      R_g[4,14] := -0.11583298;
      R_g[4,15] := 0.43668517;
      R_g[5,0] := -0.15006073;
      R_g[5,1] := 0.14857836;
      R_g[5,2] := 0.09219331;
      R_g[5,3] := 0.24307117;
      R_g[5,4] := 0.02014972;
      R_g[5,5] := -1.73904812;
      R_g[5,6] := -0.06327479;
      R_g[5,7] := 0.09475522;
      R_g[5,8] := -0.05716670;
      R_g[5,9] := 0.00648821;
      R_g[5,10] := -0.08605717;
      R_g[5,11] := 0.04396249;
      R_g[5,12] := 0.19865264;
      R_g[5,13] := 0.21015443;
      R_g[5,14] := -0.04510098;
      R_g[5,15] := -0.05707484;
      R_g[6,0] := 0.05463404;
      R_g[6,1] := -0.24671683;
      R_g[6,2] := 0.14945947;
      R_g[6,3] := 0.27781609;
      R_g[6,4] := 0.05857803;
      R_g[6,5] := -0.09827307;
      R_g[6,6] := -1.36955547;
      R_g[6,7] := 0.03997089;
      R_g[6,8] := 0.10697827;
      R_g[6,9] := -0.15282896;
      R_g[6,10] := -0.11458242;
      R_g[6,11] := 0.23231277;
      R_g[6,12] := 0.06463466;
      R_g[6,13] := -0.04114177;
      R_g[6,14] := 0.01473683;
      R_g[6,15] := 0.09800901;
      R_g[7,0] := 0.03089882;
      R_g[7,1] := -0.12866169;
      R_g[7,2] := -0.14488882;
      R_g[7,3] := 0.08099888;
      R_g[7,4] := -0.01760847;
      R_g[7,5] := 0.12323798;
      R_g[7,6] := 0.01051104;
      R_g[7,7] := -1.43148434;
      R_g[7,8] := 0.05538348;
      R_g[7,9] := 0.08765257;
      R_g[7,10] := 0.04525751;
      R_g[7,11] := -0.08530193;
      R_g[7,12] := 0.06940229;
      R_g[7,13] := 0.20471461;
      R_g[7,14] := 0.11143748;
      R_g[7,15] := -0.01617558;
      R_g[8,0] := 0.00375073;
      R_g[8,1] := 0.05561948;
      R_g[8,2] := 0.07504495;
      R_g[8,3] := 0.13846794;
      R_g[8,4] := 0.01292397;
      R_g[8,5] := -0.12762521;
      R_g[8,6] := 0.00967023;
      R_g[8,7] := -0.02755805;
      R_g[8,8] := -1.64812148;
      R_g[8,9] := 0.12763990;
      R_g[8,10] := 0.15346305;
      R_g[8,11] := -0.01111799;
      R_g[8,12] := 0.17867428;
      R_g[8,13] := -0.14499415;
      R_g[8,14] := -0.04605825;
      R_g[8,15] := 0.04006226;
      R_g[9,0] := 0.07299295;
      R_g[9,1] := -0.19717526;
      R_g[9,2] := -0.09354591;
      R_g[9,3] := 0.11423204;
      R_g[9,4] := 0.18770669;
      R_g[9,5] := -0.18770079;
      R_g[9,6] := 0.17637083;
      R_g[9,7] := -0.00016326;
      R_g[9,8] := 0.05343577;
      R_g[9,9] := -1.98581898;
      R_g[9,10] := -0.07635771;
      R_g[9,11] := 0.00779606;
      R_g[9,12] := -0.21436475;
      R_g[9,13] := 0.14591467;
      R_g[9,14] := 0.07554781;
      R_g[9,15] := -0.05975449;
      R_g[10,0] := -0.25483418;
      R_g[10,1] := 0.06535473;
      R_g[10,2] := -0.15168764;
      R_g[10,3] := -0.13676204;
      R_g[10,4] := 0.13715985;
      R_g[10,5] := -0.04971113;
      R_g[10,6] := -0.04342166;
      R_g[10,7] := 0.13203837;
      R_g[10,8] := -0.05174213;
      R_g[10,9] := 0.17224205;
      R_g[10,10] := -1.54585338;
      R_g[10,11] := 0.08824725;
      R_g[10,12] := 0.54317200;
      R_g[10,13] := -0.00582574;
      R_g[10,14] := -0.18427853;
      R_g[10,15] := -0.08446352;
      R_g[11,0] := -0.01310127;
      R_g[11,1] := 0.35428202;
      R_g[11,2] := -0.22564830;
      R_g[11,3] := -0.47703940;
      R_g[11,4] := 0.02761533;
      R_g[11,5] := -0.02962572;
      R_g[11,6] := 0.06179708;
      R_g[11,7] := -0.01533620;
      R_g[11,8] := 0.04956101;
      R_g[11,9] := 0.15626863;
      R_g[11,10] := -0.12132444;
      R_g[11,11] := -0.90700060;
      R_g[11,12] := 0.20753333;
      R_g[11,13] := -0.08345811;
      R_g[11,14] := -0.30101308;
      R_g[11,15] := -0.34388351;
      R_g[12,0] := 0.15464328;
      R_g[12,1] := -0.19553624;
      R_g[12,2] := 0.22160864;
      R_g[12,3] := 0.32764918;
      R_g[12,4] := 0.02648578;
      R_g[12,5] := 0.09656581;
      R_g[12,6] := 0.09269863;
      R_g[12,7] := -0.00748462;
      R_g[12,8] := 0.23840839;
      R_g[12,9] := -0.22269231;
      R_g[12,10] := -0.14327462;
      R_g[12,11] := 0.16783834;
      R_g[12,12] := -1.56623662;
      R_g[12,13] := -0.11016289;
      R_g[12,14] := 0.14277531;
      R_g[12,15] := 0.41838351;
      R_g[13,0] := 0.08890279;
      R_g[13,1] := -0.19905017;
      R_g[13,2] := -0.01056181;
      R_g[13,3] := 0.24786228;
      R_g[13,4] := 0.07754356;
      R_g[13,5] := 0.16554046;
      R_g[13,6] := 0.26014987;
      R_g[13,7] := 0.09906179;
      R_g[13,8] := -0.00865919;
      R_g[13,9] := -0.30192977;
      R_g[13,10] := -0.02393581;
      R_g[13,11] := -0.07343359;
      R_g[13,12] := -0.12892069;
      R_g[13,13] := -1.64273596;
      R_g[13,14] := 0.06043187;
      R_g[13,15] := 0.12883589;
      R_g[14,0] := -0.09330796;
      R_g[14,1] := 0.19971547;
      R_g[14,2] := -0.16603884;
      R_g[14,3] := -0.24762461;
      R_g[14,4] := -0.24546199;
      R_g[14,5] := -0.23372373;
      R_g[14,6] := -0.02659419;
      R_g[14,7] := 0.10576805;
      R_g[14,8] := -0.06399340;
      R_g[14,9] := 0.20369950;
      R_g[14,10] := 0.02550231;
      R_g[14,11] := -0.13061593;
      R_g[14,12] := 0.01752861;
      R_g[14,13] := -0.16408648;
      R_g[14,14] := -0.94703943;
      R_g[14,15] := -0.04546883;
      R_g[15,0] := 0.06223761;
      R_g[15,1] := 0.25574595;
      R_g[15,2] := -0.12919725;
      R_g[15,3] := -0.24720787;
      R_g[15,4] := -0.08847310;
      R_g[15,5] := 0.09416921;
      R_g[15,6] := 0.13703704;
      R_g[15,7] := 0.01633993;
      R_g[15,8] := -0.00774476;
      R_g[15,9] := 0.14204754;
      R_g[15,10] := -0.01668179;
      R_g[15,11] := -0.24296039;
      R_g[15,12] := -0.17473798;
      R_g[15,13] := -0.20718963;
      R_g[15,14] := -0.19613318;
      R_g[15,15] := -1.75475442;
      R_o[0,0] := 0.23086470;
      R_o[0,1] := -1.33466291;
      R_o[0,2] := 0.40422425;
      R_o[0,3] := 1.00496864;
      R_o[0,4] := -0.45047671;
      R_o[0,5] := 0.41842493;
      R_o[0,6] := 0.33340541;
      R_o[0,7] := 0.16748093;
      R_o[0,8] := 0.45315337;
      R_o[0,9] := -0.09557626;
      R_o[0,10] := 0.29309452;
      R_o[0,11] := -1.10283887;
      R_o[0,12] := -0.66500819;
      R_o[0,13] := -0.10580891;
      R_o[0,14] := 0.25909087;
      R_o[0,15] := 0.36167490;
      R_o[1,0] := 1.00252807;
      R_o[1,1] := -1.37035978;
      R_o[1,2] := 0.19543879;
      R_o[1,3] := 0.60937399;
      R_o[1,4] := -0.58943295;
      R_o[1,5] := 0.58583379;
      R_o[1,6] := -0.09563978;
      R_o[1,7] := 0.21723722;
      R_o[1,8] := 0.63898450;
      R_o[1,9] := 0.46265250;
      R_o[1,10] := -0.08759028;
      R_o[1,11] := -0.10910024;
      R_o[1,12] := -0.56959164;
      R_o[1,13] := -0.19031867;
      R_o[1,14] := 0.52084339;
      R_o[1,15] := -0.19041286;
      R_o[2,0] := 0.62921733;
      R_o[2,1] := -1.09719419;
      R_o[2,2] := 0.72180182;
      R_o[2,3] := 0.89839655;
      R_o[2,4] := -0.10379701;
      R_o[2,5] := 0.04743656;
      R_o[2,6] := 0.27034393;
      R_o[2,7] := -0.02836194;
      R_o[2,8] := 0.27866253;
      R_o[2,9] := -0.22055538;
      R_o[2,10] := 0.02680908;
      R_o[2,11] := -0.52208543;
      R_o[2,12] := 0.08205704;
      R_o[2,13] := -0.75110227;
      R_o[2,14] := 0.44837156;
      R_o[2,15] := 0.19737180;
      R_o[3,0] := 0.07306311;
      R_o[3,1] := -0.41626626;
      R_o[3,2] := 0.06146695;
      R_o[3,3] := -0.13822801;
      R_o[3,4] := -0.18535224;
      R_o[3,5] := 0.13184804;
      R_o[3,6] := 0.48923409;
      R_o[3,7] := 0.10094553;
      R_o[3,8] := -0.12129596;
      R_o[3,9] := 0.16955170;
      R_o[3,10] := 0.10794428;
      R_o[3,11] := -0.40550727;
      R_o[3,12] := -0.01614563;
      R_o[3,13] := -0.00363492;
      R_o[3,14] := 0.34145111;
      R_o[3,15] := -0.30746472;
      R_o[4,0] := 0.49981391;
      R_o[4,1] := -0.44877273;
      R_o[4,2] := 0.02899466;
      R_o[4,3] := 0.28911862;
      R_o[4,4] := -0.54706609;
      R_o[4,5] := 0.45331240;
      R_o[4,6] := 0.31260601;
      R_o[4,7] := 0.21592355;
      R_o[4,8] := -0.18226579;
      R_o[4,9] := -0.08202437;
      R_o[4,10] := 0.19890244;
      R_o[4,11] := -0.44599697;
      R_o[4,12] := -0.00842409;
      R_o[4,13] := 0.31605095;
      R_o[4,14] := 0.19491857;
      R_o[4,15] := 0.15177047;
      R_o[5,0] := 0.16722851;
      R_o[5,1] := -0.90651047;
      R_o[5,2] := -0.09893818;
      R_o[5,3] := 0.57212383;
      R_o[5,4] := -0.52560890;
      R_o[5,5] := 0.09904512;
      R_o[5,6] := -0.07018632;
      R_o[5,7] := 0.39063781;
      R_o[5,8] := 0.46648788;
      R_o[5,9] := -0.14858934;
      R_o[5,10] := 0.18397059;
      R_o[5,11] := -0.73446417;
      R_o[5,12] := -0.48227623;
      R_o[5,13] := 0.11307760;
      R_o[5,14] := 0.02705877;
      R_o[5,15] := -0.05367837;
      R_o[6,0] := 0.46423894;
      R_o[6,1] := -1.16708338;
      R_o[6,2] := -0.04188760;
      R_o[6,3] := 0.31886110;
      R_o[6,4] := -0.09108678;
      R_o[6,5] := -0.06297291;
      R_o[6,6] := 1.53958011;
      R_o[6,7] := -0.62613803;
      R_o[6,8] := 0.44990379;
      R_o[6,9] := -0.72628647;
      R_o[6,10] := 0.38245559;
      R_o[6,11] := -0.53905845;
      R_o[6,12] := -0.71751851;
      R_o[6,13] := 0.50797898;
      R_o[6,14] := -0.32370299;
      R_o[6,15] := -0.09905253;
      R_o[7,0] := 0.29057696;
      R_o[7,1] := -1.98383927;
      R_o[7,2] := 0.13180807;
      R_o[7,3] := 0.91098952;
      R_o[7,4] := -0.17648123;
      R_o[7,5] := 0.84703767;
      R_o[7,6] := 0.33756742;
      R_o[7,7] := 0.43434864;
      R_o[7,8] := 0.69060326;
      R_o[7,9] := 0.22266115;
      R_o[7,10] := 0.27353692;
      R_o[7,11] := -0.72814274;
      R_o[7,12] := -0.43481529;
      R_o[7,13] := 0.07530996;
      R_o[7,14] := 0.07590891;
      R_o[7,15] := 0.53633690;
      R_o[8,0] := 0.13431163;
      R_o[8,1] := -0.85810894;
      R_o[8,2] := 0.02636042;
      R_o[8,3] := 0.89655668;
      R_o[8,4] := -0.58121395;
      R_o[8,5] := 0.16582070;
      R_o[8,6] := 0.39200631;
      R_o[8,7] := 0.48816058;
      R_o[8,8] := -0.40269989;
      R_o[8,9] := -0.12494008;
      R_o[8,10] := -0.18525635;
      R_o[8,11] := -0.58216965;
      R_o[8,12] := -0.17224526;
      R_o[8,13] := -0.06991822;
      R_o[8,14] := 0.44399384;
      R_o[8,15] := 0.06420073;
      R_o[9,0] := 0.65809155;
      R_o[9,1] := -0.74305850;
      R_o[9,2] := 0.04991319;
      R_o[9,3] := 0.72979444;
      R_o[9,4] := -0.12074757;
      R_o[9,5] := -0.12410212;
      R_o[9,6] := 0.20973517;
      R_o[9,7] := 0.61132842;
      R_o[9,8] := 0.64282608;
      R_o[9,9] := -1.04169548;
      R_o[9,10] := -1.02774072;
      R_o[9,11] := -0.49568698;
      R_o[9,12] := -0.77422464;
      R_o[9,13] := 0.27705330;
      R_o[9,14] := 0.63361734;
      R_o[9,15] := 0.36834979;
      R_o[10,0] := 0.17629862;
      R_o[10,1] := -0.81763780;
      R_o[10,2] := -0.40000725;
      R_o[10,3] := 0.38086745;
      R_o[10,4] := -0.04421521;
      R_o[10,5] := 0.10713756;
      R_o[10,6] := 0.44333023;
      R_o[10,7] := 0.25184852;
      R_o[10,8] := 0.55721313;
      R_o[10,9] := -0.31075719;
      R_o[10,10] := -0.17523780;
      R_o[10,11] := -0.29524738;
      R_o[10,12] := -0.62744999;
      R_o[10,13] := -0.14156732;
      R_o[10,14] := 0.09456541;
      R_o[10,15] := 0.15875982;
      R_o[11,0] := 0.87462270;
      R_o[11,1] := -1.42915857;
      R_o[11,2] := 0.08348330;
      R_o[11,3] := 0.93353397;
      R_o[11,4] := -0.28696272;
      R_o[11,5] := 0.67741537;
      R_o[11,6] := 0.38184240;
      R_o[11,7] := 0.14032410;
      R_o[11,8] := 0.43739057;
      R_o[11,9] := 0.14584550;
      R_o[11,10] := 0.20533800;
      R_o[11,11] := 0.57373375;
      R_o[11,12] := -0.42474410;
      R_o[11,13] := -0.32885900;
      R_o[11,14] := 0.05512207;
      R_o[11,15] := 0.22504714;
      R_o[12,0] := -0.10892195;
      R_o[12,1] := -0.75056845;
      R_o[12,2] := -0.21053158;
      R_o[12,3] := 0.45154807;
      R_o[12,4] := -0.93503535;
      R_o[12,5] := 0.36019328;
      R_o[12,6] := 0.35020679;
      R_o[12,7] := 0.08578178;
      R_o[12,8] := 0.11221533;
      R_o[12,9] := 0.21497023;
      R_o[12,10] := 0.01753722;
      R_o[12,11] := -0.61306661;
      R_o[12,12] := -0.43410349;
      R_o[12,13] := 0.29725131;
      R_o[12,14] := 0.46178499;
      R_o[12,15] := 0.17685713;
      R_o[13,0] := 0.84386832;
      R_o[13,1] := -0.80496299;
      R_o[13,2] := 0.07475836;
      R_o[13,3] := 0.51488775;
      R_o[13,4] := -0.66752350;
      R_o[13,5] := 0.32658193;
      R_o[13,6] := 0.87158197;
      R_o[13,7] := -0.14368999;
      R_o[13,8] := 0.21309660;
      R_o[13,9] := -0.32924318;
      R_o[13,10] := 0.33622441;
      R_o[13,11] := -0.78933704;
      R_o[13,12] := -0.56442517;
      R_o[13,13] := 0.24916750;
      R_o[13,14] := 0.16380969;
      R_o[13,15] := 0.76749009;
      R_o[14,0] := 0.13153429;
      R_o[14,1] := -0.77425879;
      R_o[14,2] := -0.23358400;
      R_o[14,3] := 0.68574214;
      R_o[14,4] := -0.48119926;
      R_o[14,5] := -0.26408330;
      R_o[14,6] := 0.54169637;
      R_o[14,7] := -0.19132200;
      R_o[14,8] := 0.30803561;
      R_o[14,9] := 0.22515608;
      R_o[14,10] := -0.15176114;
      R_o[14,11] := -0.18082066;
      R_o[14,12] := -0.53965896;
      R_o[14,13] := 0.28110227;
      R_o[14,14] := 0.48795068;
      R_o[14,15] := 0.05904227;
      R_o[15,0] := 0.32206139;
      R_o[15,1] := -0.59116280;
      R_o[15,2] := 0.07525509;
      R_o[15,3] := 0.43309510;
      R_o[15,4] := -0.21452421;
      R_o[15,5] := -0.11838123;
      R_o[15,6] := 0.46171454;
      R_o[15,7] := 0.10131621;
      R_o[15,8] := 0.01249216;
      R_o[15,9] := -0.04199028;
      R_o[15,10] := 0.27042556;
      R_o[15,11] := 0.10062438;
      R_o[15,12] := -0.38477796;
      R_o[15,13] := -0.12011202;
      R_o[15,14] := 0.36958510;
      R_o[15,15] := 0.67342490;
      B_i[0] := 1.39581978;
      B_i[1] := 0.68250978;
      B_i[2] := 1.20262527;
      B_i[3] := 0.26746339;
      B_i[4] := 1.10431361;
      B_i[5] := 0.95270908;
      B_i[6] := 1.36736441;
      B_i[7] := 1.24711335;
      B_i[8] := 1.51264334;
      B_i[9] := 0.16206565;
      B_i[10] := 1.60950446;
      B_i[11] := 0.82160985;
      B_i[12] := 1.23546386;
      B_i[13] := 1.08165979;
      B_i[14] := 0.12467705;
      B_i[15] := 0.54986328;
      B_f[0] := 0.79174572;
      B_f[1] := -0.64133394;
      B_f[2] := 1.20450139;
      B_f[3] := -1.03967714;
      B_f[4] := 1.24121356;
      B_f[5] := 0.93169975;
      B_f[6] := 0.56517774;
      B_f[7] := 1.14514232;
      B_f[8] := 1.61746037;
      B_f[9] := 0.65368253;
      B_f[10] := 0.90967882;
      B_f[11] := -0.56739712;
      B_f[12] := 0.80123132;
      B_f[13] := 0.91223097;
      B_f[14] := -1.03880548;
      B_f[15] := 1.31209350;
      B_g[0] := 0.06687933;
      B_g[1] := -0.68397504;
      B_g[2] := 0.58139253;
      B_g[3] := 0.38107550;
      B_g[4] := -0.22040275;
      B_g[5] := 0.34854612;
      B_g[6] := 0.35342124;
      B_g[7] := 0.09094166;
      B_g[8] := -0.19340213;
      B_g[9] := -0.22835979;
      B_g[10] := 0.00825962;
      B_g[11] := 0.16006482;
      B_g[12] := -0.36459130;
      B_g[13] := -0.06400946;
      B_g[14] := 0.27469134;
      B_g[15] := 0.11084859;
      B_o[0] := 2.83054423;
      B_o[1] := 2.38222671;
      B_o[2] := 2.63261795;
      B_o[3] := 1.95818925;
      B_o[4] := 2.31596231;
      B_o[5] := 2.64208364;
      B_o[6] := 3.44678116;
      B_o[7] := 3.71243334;
      B_o[8] := 2.57036018;
      B_o[9] := 2.55204439;
      B_o[10] := 2.07645392;
      B_o[11] := 2.16894150;
      B_o[12] := 2.77243233;
      B_o[13] := 3.07682300;
      B_o[14] := 1.65793490;
      B_o[15] := 2.28551698;
      FC_W[0,0] := -0.53302634;
      FC_W[0,1] := 0.68295699;
      FC_W[0,2] := -0.62599581;
      FC_W[0,3] := -0.32720318;
      FC_W[0,4] := -0.08957181;
      FC_W[0,5] := -0.16555449;
      FC_W[0,6] := 0.06407359;
      FC_W[0,7] := 0.20225702;
      FC_W[0,8] := -1.04729974;
      FC_W[0,9] := -1.63024998;
      FC_W[0,10] := -0.36511818;
      FC_W[0,11] := -0.61756939;
      FC_W[0,12] := -0.26097849;
      FC_W[0,13] := 0.79630882;
      FC_W[0,14] := 0.06587959;
      FC_W[0,15] := 1.50049973;
      FC_W[1,0] := -0.11588198;
      FC_W[1,1] := 0.60197467;
      FC_W[1,2] := 0.98438090;
      FC_W[1,3] := -0.12106090;
      FC_W[1,4] := 0.36372337;
      FC_W[1,5] := 0.08963854;
      FC_W[1,6] := -1.69355536;
      FC_W[1,7] := -0.84128761;
      FC_W[1,8] := -0.09554562;
      FC_W[1,9] := -0.33927256;
      FC_W[1,10] := 1.17080462;
      FC_W[1,11] := 1.69248676;
      FC_W[1,12] := -0.02792989;
      FC_W[1,13] := 0.25264657;
      FC_W[1,14] := 1.54547310;
      FC_W[1,15] := -0.59855837;
      FC_W[2,0] := -0.56375182;
      FC_W[2,1] := 0.73003334;
      FC_W[2,2] := -0.54087758;
      FC_W[2,3] := -0.42607835;
      FC_W[2,4] := -0.14161965;
      FC_W[2,5] := -0.13632999;
      FC_W[2,6] := -0.02574298;
      FC_W[2,7] := 0.24827254;
      FC_W[2,8] := -1.09977758;
      FC_W[2,9] := -1.69800615;
      FC_W[2,10] := -0.41489336;
      FC_W[2,11] := -0.66403556;
      FC_W[2,12] := -0.25348228;
      FC_W[2,13] := 0.84585100;
      FC_W[2,14] := 0.03002551;
      FC_W[2,15] := 1.51456881;
      FC_W[3,0] := -0.19130252;
      FC_W[3,1] := 0.22978918;
      FC_W[3,2] := 0.32297230;
      FC_W[3,3] := 0.21441473;
      FC_W[3,4] := 0.31629598;
      FC_W[3,5] := -0.00644177;
      FC_W[3,6] := 0.57398194;
      FC_W[3,7] := -0.09706475;
      FC_W[3,8] := -0.05950126;
      FC_W[3,9] := -1.09413004;
      FC_W[3,10] := 0.25704047;
      FC_W[3,11] := 0.66124117;
      FC_W[3,12] := -0.31906813;
      FC_W[3,13] := 0.53711319;
      FC_W[3,14] := -1.58713961;
      FC_W[3,15] := 0.01048408;
      FC_W[4,0] := 0.31414661;
      FC_W[4,1] := -0.34332627;
      FC_W[4,2] := 0.89117354;
      FC_W[4,3] := -0.71509856;
      FC_W[4,4] := 0.09996962;
      FC_W[4,5] := -0.02766594;
      FC_W[4,6] := 0.51257795;
      FC_W[4,7] := -0.91753322;
      FC_W[4,8] := 1.08904767;
      FC_W[4,9] := -0.05996554;
      FC_W[4,10] := -1.12754261;
      FC_W[4,11] := -0.16949877;
      FC_W[4,12] := -0.76937914;
      FC_W[4,13] := -1.22835076;
      FC_W[4,14] := -0.38305089;
      FC_W[4,15] := 1.15847588;
      FC_W[5,0] := 0.66654950;
      FC_W[5,1] := -0.55389386;
      FC_W[5,2] := -1.28292799;
      FC_W[5,3] := 0.23086897;
      FC_W[5,4] := -0.46505886;
      FC_W[5,5] := -2.09175372;
      FC_W[5,6] := -0.96113479;
      FC_W[5,7] := 1.04218686;
      FC_W[5,8] := 1.51852155;
      FC_W[5,9] := -3.80393577;
      FC_W[5,10] := -1.47868264;
      FC_W[5,11] := -0.25626692;
      FC_W[5,12] := 0.24388616;
      FC_W[5,13] := 0.11551145;
      FC_W[5,14] := -0.36641932;
      FC_W[5,15] := -1.08498335;
      FC_W[6,0] := 0.43836260;
      FC_W[6,1] := 0.89048672;
      FC_W[6,2] := 0.11603133;
      FC_W[6,3] := 0.96929032;
      FC_W[6,4] := 1.08512294;
      FC_W[6,5] := -0.51023304;
      FC_W[6,6] := -0.43371543;
      FC_W[6,7] := 1.29686451;
      FC_W[6,8] := -0.10809528;
      FC_W[6,9] := -0.04550074;
      FC_W[6,10] := -0.73365164;
      FC_W[6,11] := 0.29729211;
      FC_W[6,12] := -0.41153616;
      FC_W[6,13] := -0.01893469;
      FC_W[6,14] := -0.83904946;
      FC_W[6,15] := -0.24609792;
      FC_W[7,0] := -0.18477769;
      FC_W[7,1] := 0.20369241;
      FC_W[7,2] := 0.28273052;
      FC_W[7,3] := 0.25776774;
      FC_W[7,4] := 0.33915454;
      FC_W[7,5] := -0.02453313;
      FC_W[7,6] := 0.63038129;
      FC_W[7,7] := -0.08684690;
      FC_W[7,8] := -0.03923411;
      FC_W[7,9] := -1.06299269;
      FC_W[7,10] := 0.25988910;
      FC_W[7,11] := 0.64730209;
      FC_W[7,12] := -0.33632410;
      FC_W[7,13] := 0.53152817;
      FC_W[7,14] := -1.56968188;
      FC_W[7,15] := 0.01425198;
      FC_W[8,0] := -0.21285072;
      FC_W[8,1] := 0.28717902;
      FC_W[8,2] := 0.31703505;
      FC_W[8,3] := 0.15400071;
      FC_W[8,4] := 0.33542806;
      FC_W[8,5] := -0.01905481;
      FC_W[8,6] := 0.53315622;
      FC_W[8,7] := -0.09981918;
      FC_W[8,8] := -0.08895166;
      FC_W[8,9] := -1.12627339;
      FC_W[8,10] := 0.25810486;
      FC_W[8,11] := 0.67377931;
      FC_W[8,12] := -0.26128903;
      FC_W[8,13] := 0.54103297;
      FC_W[8,14] := -1.60691571;
      FC_W[8,15] := -0.01362194;
      FC_W[9,0] := -0.19543010;
      FC_W[9,1] := 0.21304309;
      FC_W[9,2] := 0.29270205;
      FC_W[9,3] := 0.23064727;
      FC_W[9,4] := 0.32767618;
      FC_W[9,5] := -0.02455352;
      FC_W[9,6] := 0.59843177;
      FC_W[9,7] := -0.08202294;
      FC_W[9,8] := -0.06203229;
      FC_W[9,9] := -1.09027541;
      FC_W[9,10] := 0.26965019;
      FC_W[9,11] := 0.65412533;
      FC_W[9,12] := -0.33295867;
      FC_W[9,13] := 0.54472339;
      FC_W[9,14] := -1.58246577;
      FC_W[9,15] := 0.00871467;
      FC_W[10,0] := -0.44877350;
      FC_W[10,1] := -0.27872828;
      FC_W[10,2] := -0.20872270;
      FC_W[10,3] := -0.59951437;
      FC_W[10,4] := -0.64611596;
      FC_W[10,5] := -0.55243987;
      FC_W[10,6] := 0.24780296;
      FC_W[10,7] := -0.74007368;
      FC_W[10,8] := 0.32341728;
      FC_W[10,9] := -2.57707667;
      FC_W[10,10] := 0.57498157;
      FC_W[10,11] := 0.61854416;
      FC_W[10,12] := 0.01876899;
      FC_W[10,13] := 0.75633305;
      FC_W[10,14] := -0.89730561;
      FC_W[10,15] := -0.39787960;
      FC_W[11,0] := 0.61467212;
      FC_W[11,1] := 0.19168422;
      FC_W[11,2] := 0.93443829;
      FC_W[11,3] := -0.59301579;
      FC_W[11,4] := -0.92330587;
      FC_W[11,5] := 0.40248036;
      FC_W[11,6] := 0.63603044;
      FC_W[11,7] := 0.38971198;
      FC_W[11,8] := -0.51435661;
      FC_W[11,9] := -0.25507462;
      FC_W[11,10] := -0.58355647;
      FC_W[11,11] := 0.01116155;
      FC_W[11,12] := -1.25048304;
      FC_W[11,13] := -0.29360211;
      FC_W[11,14] := 0.33364284;
      FC_W[11,15] := -1.04067647;
      FC_W[12,0] := 0.22212029;
      FC_W[12,1] := -0.14197727;
      FC_W[12,2] := 1.13170397;
      FC_W[12,3] := -0.61373824;
      FC_W[12,4] := -0.75162232;
      FC_W[12,5] := 0.45277873;
      FC_W[12,6] := 0.43703261;
      FC_W[12,7] := 0.68883568;
      FC_W[12,8] := -0.27114886;
      FC_W[12,9] := -0.33246922;
      FC_W[12,10] := -0.36722985;
      FC_W[12,11] := -0.21226645;
      FC_W[12,12] := -1.38135302;
      FC_W[12,13] := -0.28390571;
      FC_W[12,14] := 0.21292266;
      FC_W[12,15] := -1.02846980;
      FC_W[13,0] := -0.42784557;
      FC_W[13,1] := -1.55966008;
      FC_W[13,2] := -0.23814020;
      FC_W[13,3] := 0.81332529;
      FC_W[13,4] := 1.01786804;
      FC_W[13,5] := -0.76350653;
      FC_W[13,6] := 0.04761689;
      FC_W[13,7] := -0.52871329;
      FC_W[13,8] := -0.08105175;
      FC_W[13,9] := -0.55568081;
      FC_W[13,10] := 1.00466228;
      FC_W[13,11] := 1.32452846;
      FC_W[13,12] := -1.16723299;
      FC_W[13,13] := 1.34940958;
      FC_W[13,14] := 2.63829517;
      FC_W[13,15] := -0.22661680;
      FC_W[14,0] := -2.35853815;
      FC_W[14,1] := 0.42897072;
      FC_W[14,2] := -1.65632534;
      FC_W[14,3] := -1.45689034;
      FC_W[14,4] := -0.23707533;
      FC_W[14,5] := 2.00690389;
      FC_W[14,6] := 1.07422280;
      FC_W[14,7] := 2.12480640;
      FC_W[14,8] := 1.78673518;
      FC_W[14,9] := 0.14402351;
      FC_W[14,10] := -1.98161817;
      FC_W[14,11] := 2.80044842;
      FC_W[14,12] := 0.03338763;
      FC_W[14,13] := 0.41240925;
      FC_W[14,14] := 1.21908247;
      FC_W[14,15] := 0.18715070;
      FC_W[15,0] := 0.94744486;
      FC_W[15,1] := 0.56090069;
      FC_W[15,2] := 0.77292573;
      FC_W[15,3] := -0.47338617;
      FC_W[15,4] := -1.32521272;
      FC_W[15,5] := 0.16259588;
      FC_W[15,6] := 0.54934692;
      FC_W[15,7] := -0.00915920;
      FC_W[15,8] := -0.71907353;
      FC_W[15,9] := -0.03908357;
      FC_W[15,10] := -0.98591125;
      FC_W[15,11] := 0.30310348;
      FC_W[15,12] := -0.98413241;
      FC_W[15,13] := 0.09539948;
      FC_W[15,14] := 0.45499024;
      FC_W[15,15] := -0.95317203;
      FC_W[16,0] := -0.90791857;
      FC_W[16,1] := 1.47015476;
      FC_W[16,2] := 1.46804285;
      FC_W[16,3] := -0.39122909;
      FC_W[16,4] := -2.34223771;
      FC_W[16,5] := -2.31965876;
      FC_W[16,6] := -0.78383219;
      FC_W[16,7] := 0.00836219;
      FC_W[16,8] := 1.98210740;
      FC_W[16,9] := 1.16555631;
      FC_W[16,10] := -1.21075189;
      FC_W[16,11] := 0.59300679;
      FC_W[16,12] := 0.61776960;
      FC_W[16,13] := 3.99444842;
      FC_W[16,14] := 0.01262518;
      FC_W[16,15] := 1.04920304;
      FC_W[17,0] := -2.79870629;
      FC_W[17,1] := -1.42033422;
      FC_W[17,2] := 1.69065225;
      FC_W[17,3] := -0.66839701;
      FC_W[17,4] := 1.27351940;
      FC_W[17,5] := 0.02801782;
      FC_W[17,6] := -0.33793277;
      FC_W[17,7] := 2.32656717;
      FC_W[17,8] := 2.14157987;
      FC_W[17,9] := -0.63859951;
      FC_W[17,10] := 1.59767425;
      FC_W[17,11] := -2.15692639;
      FC_W[17,12] := -0.74494350;
      FC_W[17,13] := 0.14399342;
      FC_W[17,14] := -0.38486624;
      FC_W[17,15] := 0.08045793;
      FC_W[18,0] := 1.34154665;
      FC_W[18,1] := 3.19789124;
      FC_W[18,2] := -1.12263572;
      FC_W[18,3] := -0.72371221;
      FC_W[18,4] := -1.43890095;
      FC_W[18,5] := 1.35449719;
      FC_W[18,6] := 1.00367022;
      FC_W[18,7] := 0.11557481;
      FC_W[18,8] := 1.42845428;
      FC_W[18,9] := -0.04815372;
      FC_W[18,10] := 1.82935095;
      FC_W[18,11] := -1.33503389;
      FC_W[18,12] := -5.11765480;
      FC_W[18,13] := -1.06049836;
      FC_W[18,14] := -0.81516898;
      FC_W[18,15] := 0.03152023;
      FC_W[19,0] := -0.15235230;
      FC_W[19,1] := -1.04747820;
      FC_W[19,2] := 1.24190295;
      FC_W[19,3] := -0.41053832;
      FC_W[19,4] := -0.26765159;
      FC_W[19,5] := 0.35931253;
      FC_W[19,6] := 0.11906569;
      FC_W[19,7] := 0.74638200;
      FC_W[19,8] := -0.61629355;
      FC_W[19,9] := -0.36762637;
      FC_W[19,10] := -0.64761603;
      FC_W[19,11] := -0.01234968;
      FC_W[19,12] := -0.39466342;
      FC_W[19,13] := -0.31511360;
      FC_W[19,14] := 0.30823269;
      FC_W[19,15] := -1.08234417;
      FC_W[20,0] := 0.26440981;
      FC_W[20,1] := -1.47835481;
      FC_W[20,2] := 0.11839479;
      FC_W[20,3] := -1.16043782;
      FC_W[20,4] := -1.16143334;
      FC_W[20,5] := 0.02869733;
      FC_W[20,6] := 0.73862082;
      FC_W[20,7] := -0.69498312;
      FC_W[20,8] := 0.40190154;
      FC_W[20,9] := -0.16530611;
      FC_W[20,10] := 0.89126289;
      FC_W[20,11] := 0.34054285;
      FC_W[20,12] := -0.26115537;
      FC_W[20,13] := -0.38540450;
      FC_W[20,14] := 0.68782163;
      FC_W[20,15] := 0.64379901;
      FC_W[21,0] := -0.66346151;
      FC_W[21,1] := 0.58732224;
      FC_W[21,2] := 0.06739193;
      FC_W[21,3] := 0.97263134;
      FC_W[21,4] := -0.86781269;
      FC_W[21,5] := -1.02743030;
      FC_W[21,6] := 0.16887170;
      FC_W[21,7] := 1.69680274;
      FC_W[21,8] := -1.14409292;
      FC_W[21,9] := 0.14942116;
      FC_W[21,10] := 0.32693279;
      FC_W[21,11] := 0.61105758;
      FC_W[21,12] := 0.16232388;
      FC_W[21,13] := -1.26744127;
      FC_W[21,14] := -0.87755442;
      FC_W[21,15] := 0.54278499;
      FC_W[22,0] := 0.28525919;
      FC_W[22,1] := -1.50926864;
      FC_W[22,2] := 1.53992140;
      FC_W[22,3] := 1.62703526;
      FC_W[22,4] := -0.20404652;
      FC_W[22,5] := 0.43128183;
      FC_W[22,6] := -0.04736441;
      FC_W[22,7] := 0.18942423;
      FC_W[22,8] := 0.26407915;
      FC_W[22,9] := -0.95513147;
      FC_W[22,10] := -0.04719095;
      FC_W[22,11] := 1.31737375;
      FC_W[22,12] := -0.56206286;
      FC_W[22,13] := -0.34498781;
      FC_W[22,14] := 1.28337383;
      FC_W[22,15] := 1.78748143;
      FC_W[23,0] := -0.06120704;
      FC_W[23,1] := -1.64042079;
      FC_W[23,2] := -0.25326556;
      FC_W[23,3] := 1.11953604;
      FC_W[23,4] := 1.08679652;
      FC_W[23,5] := -0.38698131;
      FC_W[23,6] := 0.44496018;
      FC_W[23,7] := -0.78417253;
      FC_W[23,8] := 0.07545953;
      FC_W[23,9] := -0.68813795;
      FC_W[23,10] := 0.98399347;
      FC_W[23,11] := 1.54028356;
      FC_W[23,12] := -1.13344729;
      FC_W[23,13] := 1.85424924;
      FC_W[23,14] := 2.03626943;
      FC_W[23,15] := -0.30457237;
      FC_W[24,0] := 0.22877936;
      FC_W[24,1] := -1.47323406;
      FC_W[24,2] := 1.46277165;
      FC_W[24,3] := 1.76430011;
      FC_W[24,4] := -0.24940053;
      FC_W[24,5] := 0.43059126;
      FC_W[24,6] := 0.07592186;
      FC_W[24,7] := 0.14821550;
      FC_W[24,8] := 0.34645149;
      FC_W[24,9] := -0.87015730;
      FC_W[24,10] := -0.04559883;
      FC_W[24,11] := 1.23906600;
      FC_W[24,12] := -0.71117419;
      FC_W[24,13] := -0.41323856;
      FC_W[24,14] := 1.30650675;
      FC_W[24,15] := 1.71300721;
      FC_W[25,0] := 0.22861326;
      FC_W[25,1] := -1.47545123;
      FC_W[25,2] := 1.46235204;
      FC_W[25,3] := 1.76556575;
      FC_W[25,4] := -0.24908429;
      FC_W[25,5] := 0.43040714;
      FC_W[25,6] := 0.07507181;
      FC_W[25,7] := 0.14740342;
      FC_W[25,8] := 0.34566393;
      FC_W[25,9] := -0.86833739;
      FC_W[25,10] := -0.04680423;
      FC_W[25,11] := 1.23651314;
      FC_W[25,12] := -0.70846480;
      FC_W[25,13] := -0.41374815;
      FC_W[25,14] := 1.30441546;
      FC_W[25,15] := 1.71272981;
      FC_W[26,0] := 0.38304979;
      FC_W[26,1] := -1.76469123;
      FC_W[26,2] := 1.27260387;
      FC_W[26,3] := 0.61524868;
      FC_W[26,4] := 0.92497736;
      FC_W[26,5] := 0.40269154;
      FC_W[26,6] := -0.54810572;
      FC_W[26,7] := -0.81347013;
      FC_W[26,8] := 0.52034670;
      FC_W[26,9] := -0.98628432;
      FC_W[26,10] := -0.39365792;
      FC_W[26,11] := 1.14341772;
      FC_W[26,12] := 0.13778362;
      FC_W[26,13] := 0.94409907;
      FC_W[26,14] := 1.57374060;
      FC_W[26,15] := 0.79883248;
      FC_W[27,0] := -1.14280367;
      FC_W[27,1] := 0.59307718;
      FC_W[27,2] := -0.26207438;
      FC_W[27,3] := 0.87626535;
      FC_W[27,4] := -0.93659830;
      FC_W[27,5] := -1.49864197;
      FC_W[27,6] := 0.44960785;
      FC_W[27,7] := 1.37962472;
      FC_W[27,8] := -1.18801665;
      FC_W[27,9] := 0.41698411;
      FC_W[27,10] := 0.34206629;
      FC_W[27,11] := 0.51468468;
      FC_W[27,12] := 0.28827220;
      FC_W[27,13] := -1.38293719;
      FC_W[27,14] := -1.01115930;
      FC_W[27,15] := 0.12471072;
      FC_W[28,0] := 0.04424974;
      FC_W[28,1] := 0.13536097;
      FC_W[28,2] := 0.75559741;
      FC_W[28,3] := -0.35790223;
      FC_W[28,4] := 1.36025250;
      FC_W[28,5] := -0.88536996;
      FC_W[28,6] := -0.00372644;
      FC_W[28,7] := -0.29969507;
      FC_W[28,8] := 0.19030553;
      FC_W[28,9] := -0.01632601;
      FC_W[28,10] := -1.65227020;
      FC_W[28,11] := 0.34139770;
      FC_W[28,12] := -0.34939787;
      FC_W[28,13] := -0.57886147;
      FC_W[28,14] := -0.35904202;
      FC_W[28,15] := 0.34676898;
      FC_W[29,0] := -0.38553143;
      FC_W[29,1] := 1.27834022;
      FC_W[29,2] := -1.67743385;
      FC_W[29,3] := -1.05788505;
      FC_W[29,4] := 0.22803551;
      FC_W[29,5] := -0.11723094;
      FC_W[29,6] := 0.36204663;
      FC_W[29,7] := -0.44841900;
      FC_W[29,8] := 0.03538510;
      FC_W[29,9] := 1.20318663;
      FC_W[29,10] := -0.20551582;
      FC_W[29,11] := -1.71424949;
      FC_W[29,12] := 0.49145132;
      FC_W[29,13] := 0.40932351;
      FC_W[29,14] := -1.01760292;
      FC_W[29,15] := -1.91052508;
      FC_W[30,0] := 0.28723446;
      FC_W[30,1] := -1.51120055;
      FC_W[30,2] := 1.54199433;
      FC_W[30,3] := 1.62217951;
      FC_W[30,4] := -0.20229872;
      FC_W[30,5] := 0.43358997;
      FC_W[30,6] := -0.05039101;
      FC_W[30,7] := 0.18811959;
      FC_W[30,8] := 0.26187438;
      FC_W[30,9] := -0.95781857;
      FC_W[30,10] := -0.04945299;
      FC_W[30,11] := 1.31731784;
      FC_W[30,12] := -0.55758446;
      FC_W[30,13] := -0.34352461;
      FC_W[30,14] := 1.28357959;
      FC_W[30,15] := 1.78932595;
      FC_W[31,0] := 0.33338901;
      FC_W[31,1] := -1.51106906;
      FC_W[31,2] := 1.56730652;
      FC_W[31,3] := 1.55137372;
      FC_W[31,4] := -0.17190555;
      FC_W[31,5] := 0.45433214;
      FC_W[31,6] := -0.09396910;
      FC_W[31,7] := 0.22680379;
      FC_W[31,8] := 0.23822255;
      FC_W[31,9] := -0.98215002;
      FC_W[31,10] := -0.06985018;
      FC_W[31,11] := 1.32410133;
      FC_W[31,12] := -0.49385709;
      FC_W[31,13] := -0.31897312;
      FC_W[31,14] := 1.26462150;
      FC_W[31,15] := 1.82302165;
      FC_W[32,0] := 0.22924727;
      FC_W[32,1] := -1.46797276;
      FC_W[32,2] := 1.56526399;
      FC_W[32,3] := 1.58788276;
      FC_W[32,4] := -0.22412077;
      FC_W[32,5] := 0.25628337;
      FC_W[32,6] := -0.05829662;
      FC_W[32,7] := 0.24949729;
      FC_W[32,8] := 0.18913403;
      FC_W[32,9] := -0.95914072;
      FC_W[32,10] := -0.00602742;
      FC_W[32,11] := 1.44420707;
      FC_W[32,12] := -0.56866109;
      FC_W[32,13] := -0.45418915;
      FC_W[32,14] := 1.21856201;
      FC_W[32,15] := 1.79085994;
      FC_W[33,0] := 0.27113631;
      FC_W[33,1] := -1.44990373;
      FC_W[33,2] := 1.67819250;
      FC_W[33,3] := 1.38159657;
      FC_W[33,4] := -0.19107535;
      FC_W[33,5] := 0.18168713;
      FC_W[33,6] := -0.21811114;
      FC_W[33,7] := 0.35240412;
      FC_W[33,8] := 0.06086530;
      FC_W[33,9] := -1.05922282;
      FC_W[33,10] := -0.01789864;
      FC_W[33,11] := 1.57391202;
      FC_W[33,12] := -0.37516510;
      FC_W[33,13] := -0.46472317;
      FC_W[33,14] := 1.11760533;
      FC_W[33,15] := 1.88658249;
      FC_W[34,0] := 0.32269877;
      FC_W[34,1] := -1.43542671;
      FC_W[34,2] := 1.66118479;
      FC_W[34,3] := 1.39128089;
      FC_W[34,4] := -0.20390645;
      FC_W[34,5] := 0.26313210;
      FC_W[34,6] := -0.20318714;
      FC_W[34,7] := 0.32080358;
      FC_W[34,8] := 0.10883178;
      FC_W[34,9] := -1.06268609;
      FC_W[34,10] := -0.01133159;
      FC_W[34,11] := 1.51307917;
      FC_W[34,12] := -0.43998954;
      FC_W[34,13] := -0.41575021;
      FC_W[34,14] := 1.14673424;
      FC_W[34,15] := 1.89976144;
      FC_W[35,0] := 0.18407848;
      FC_W[35,1] := -1.46272326;
      FC_W[35,2] := 1.47307324;
      FC_W[35,3] := 1.66796565;
      FC_W[35,4] := -0.24057212;
      FC_W[35,5] := 0.21155888;
      FC_W[35,6] := 0.05332418;
      FC_W[35,7] := 0.21069987;
      FC_W[35,8] := 0.23600885;
      FC_W[35,9] := -0.89149302;
      FC_W[35,10] := 0.04807700;
      FC_W[35,11] := 1.42777205;
      FC_W[35,12] := -0.71111673;
      FC_W[35,13] := -0.46023691;
      FC_W[35,14] := 1.25808752;
      FC_W[35,15] := 1.70261586;
      FC_W[36,0] := -2.86385798;
      FC_W[36,1] := -0.52148002;
      FC_W[36,2] := -0.29675904;
      FC_W[36,3] := 4.63355112;
      FC_W[36,4] := -1.54004574;
      FC_W[36,5] := 0.87013870;
      FC_W[36,6] := 1.44518447;
      FC_W[36,7] := -2.18261647;
      FC_W[36,8] := 0.82160705;
      FC_W[36,9] := -0.17502466;
      FC_W[36,10] := -0.96307951;
      FC_W[36,11] := -1.56679106;
      FC_W[36,12] := -0.41614529;
      FC_W[36,13] := -0.69842845;
      FC_W[36,14] := 1.35561681;
      FC_W[36,15] := -0.05721238;
      FC_W[37,0] := 0.15488347;
      FC_W[37,1] := -1.45589542;
      FC_W[37,2] := 1.44418216;
      FC_W[37,3] := 1.71133900;
      FC_W[37,4] := -0.24417210;
      FC_W[37,5] := 0.19820066;
      FC_W[37,6] := 0.08134115;
      FC_W[37,7] := 0.19478567;
      FC_W[37,8] := 0.24365275;
      FC_W[37,9] := -0.87144059;
      FC_W[37,10] := 0.05783046;
      FC_W[37,11] := 1.41966331;
      FC_W[37,12] := -0.74120307;
      FC_W[37,13] := -0.45803425;
      FC_W[37,14] := 1.27259934;
      FC_W[37,15] := 1.66730762;
      FC_W[38,0] := -0.21534352;
      FC_W[38,1] := -1.96326339;
      FC_W[38,2] := -0.75508815;
      FC_W[38,3] := 1.20778084;
      FC_W[38,4] := -1.46449494;
      FC_W[38,5] := -0.21948476;
      FC_W[38,6] := -3.29061508;
      FC_W[38,7] := -0.74855620;
      FC_W[38,8] := 0.25157410;
      FC_W[38,9] := 1.20771646;
      FC_W[38,10] := -0.30755150;
      FC_W[38,11] := 0.98883963;
      FC_W[38,12] := -0.96645385;
      FC_W[38,13] := 1.24448228;
      FC_W[38,14] := -2.63472676;
      FC_W[38,15] := 1.38428092;
      FC_W[39,0] := -1.46080005;
      FC_W[39,1] := -0.90218180;
      FC_W[39,2] := -1.38880670;
      FC_W[39,3] := -0.08306644;
      FC_W[39,4] := -0.66849297;
      FC_W[39,5] := 1.32543874;
      FC_W[39,6] := -1.17536473;
      FC_W[39,7] := 0.81609625;
      FC_W[39,8] := 1.06732941;
      FC_W[39,9] := 0.58146608;
      FC_W[39,10] := -1.25798881;
      FC_W[39,11] := 2.07855940;
      FC_W[39,12] := -0.38577294;
      FC_W[39,13] := 0.62384450;
      FC_W[39,14] := -0.81358123;
      FC_W[39,15] := 0.89604688;
      FC_B[0] := 0.02629896;
      FC_B[1] := 0.42752317;
      FC_B[2] := 0.01502107;
      FC_B[3] := -0.10187675;
      FC_B[4] := -0.33405676;
      FC_B[5] := 0.41800657;
      FC_B[6] := 0.26909930;
      FC_B[7] := -0.10668041;
      FC_B[8] := -0.05807845;
      FC_B[9] := -0.10296487;
      FC_B[10] := 0.06830941;
      FC_B[11] := -0.82022250;
      FC_B[12] := -0.82363302;
      FC_B[13] := -0.48747486;
      FC_B[14] := 0.40635556;
      FC_B[15] := -0.74980736;
      FC_B[16] := 0.52938378;
      FC_B[17] := -0.02519251;
      FC_B[18] := 0.72231776;
      FC_B[19] := -0.97234488;
      FC_B[20] := -0.66601145;
      FC_B[21] := 0.17456011;
      FC_B[22] := -1.32404578;
      FC_B[23] := -0.70627439;
      FC_B[24] := -1.30787647;
      FC_B[25] := -1.30782068;
      FC_B[26] := -1.02975488;
      FC_B[27] := 0.43721533;
      FC_B[28] := 0.05014376;
      FC_B[29] := 1.18653333;
      FC_B[30] := -1.32503390;
      FC_B[31] := -1.32861042;
      FC_B[32] := -1.27917075;
      FC_B[33] := -1.26075757;
      FC_B[34] := -1.27981257;
      FC_B[35] := -1.26051843;
      FC_B[36] := -0.34180054;
      FC_B[37] := -1.24986994;
      FC_B[38] := 0.50247991;
      FC_B[39] := 0.46928239;

END_DATA_BLOCK
